Universal Robots URScript: PgProg.script

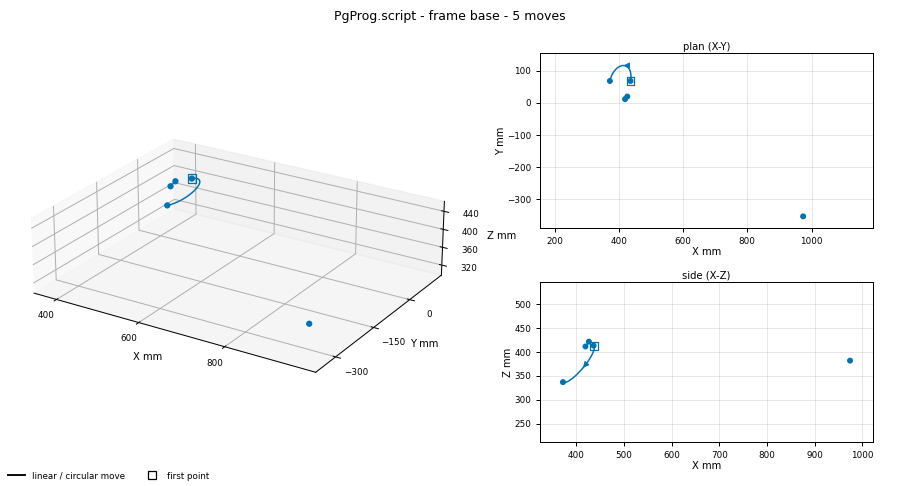
[picture p0: tool path of PgProg.script in frame base, 5 of 9 moves have a stored position in this frame; points joined in program order, loops and branches not executed]
def PgProg():
  # Global parameters:
  global speed_ms    = 0.250
  global speed_rads  = 0.750
  global accel_mss   = 1.200
  global accel_radss = 1.200
  global blend_radius_m = 0.000

  #--------------------------
  # Add any default subprograms here
  # For example, to drive a gripper as a program call:
  # def Gripper_Open():
  #   ...
  # end
  #
  # Example to drive a spray gun:
  def SprayOn(value):
    # use the value as an output:
    DO_SPRAY = 5
    if value == 0:
      set_standard_digital_out(DO_SPRAY, False)
    else:
      set_standard_digital_out(DO_SPRAY, True)
    end
  end

  # Example to synchronize 2
  def Synchronize():
    # Use the following digital output to signal the state of the robot:
    DO_SYNC = 1

    # Use the following digital input to get the state of another robot:
    DI_SYNC = 1

    if (get_standard_digital_out(DO_SYNC) == get_standard_digital_in(DI_SYNC)):
      set_standard_digital_out(DO_SYNC, not (get_standard_digital_out(DI_SYNC)))
      sleep(0.1)
      thread Thread_wait_1():
        while (True):
          sleep(0.01)
        end
      end
      if (get_standard_digital_out(DO_SYNC) != get_standard_digital_in(DI_SYNC)):
        global thread_handler_1=run Thread_wait_1()
        while (get_standard_digital_out(DO_SYNC) != get_standard_digital_in(DI_SYNC)):
          sync()
        end
        kill thread_handler_1
      end
    else:
      if (get_standard_digital_out(DO_SYNC) != get_standard_digital_in(DI_SYNC)):
        set_standard_digital_out(DO_SYNC, not (get_standard_digital_out(DO_SYNC)))
      end
    end
  end

  #
  # Example to move an external axis
  def MoveAxis(value):
    # use the value as an output:
    DO_AXIS_1 = 1
    DI_AXIS_1 = 1
    if value <= 0:
      set_standard_digital_out(DO_AXIS_1, False)

      # Wait for digital input to change state
      #while (get_standard_digital_in(DI_AXIS_1) != False):
      #  sync()
      #end
    else:
      set_standard_digital_out(DO_AXIS_1, True)

      # Wait for digital input to change state
      #while (get_standard_digital_in(DI_AXIS_1) != True):
      #  sync()
      #end
    end
  end
  #--------------------------


  # Main program:
  # Program generated by RoboDK v6.0.7 for ABB IRB 120-3/0.6 on XX/XX/XXXX 18:00:00
  # Using nominal kinematics.
  # Using Ref. Frame Pg: p[1.234570, -0.098765, 0.050500, 0.000000, 0.000000, 0.523599]
  # set_reference(p[1.234570, -0.098765, 0.050500, 0.000000, 0.000000, 0.523599])
  # Using TCP Tool Pg: p[0.010000, 0.020000, 0.150000, 0.261799, 0.000000, 0.000000]
  set_tcp(p[0.010000, 0.020000, 0.150000, 0.261799, 0.000000, 0.000000])
  speed_ms    = 0.2500
  blend_radius_m = 0.0050
  movej([0.000000, -0.174533, 0.349066, 0.000000, 0.523599, 0.000000],1.20000,0.75000,0,0.0000)
  movel(p[0.436232, 0.068297, 0.413715, 0.138328, 2.253250, -0.296646],accel_mss,speed_ms,0,0.005)
  # Circular move (R50.0 mm)
  movec(p[0.414005, 0.116593, 0.367095, 0.138328, 2.253250, -0.296646],p[0.371953, 0.068296, 0.337111, 0.138328, 2.253250, -0.296646],1.20000,0.25000,0.0050)
  movej([0.349066, -0.174533, 0.349066, 0.000000, 0.523599, 0.000000],1.20000,0.75000,0,0.0000)
  accel_radss = 2.094
  speed_rads  = 1.0472
  accel_mss   = 0.8000
  speed_ms    = 0.1000
  movel(p[0.419189, 0.011793, 0.411899, 0.138328, 2.253250, -0.296646],accel_mss,speed_ms,0,0.000)
  blend_radius_m = 0.0000
  movel(p[0.426318, 0.020000, 0.422034, 0.138328, 2.253250, -0.296646],accel_mss,speed_ms,0,0.000)
  sleep(0.500)
  halt() # reimplement this function to force stop
  popup("Hello from postgen","Message",False,False,blocking=True)
  # a comment
  SubProgram()
  CustomCode(42)
  ThreadProg
  set_standard_digital_out(1, True)
  Valve = False
  set_standard_digital_out(3, 2.5)
  while (get_standard_digital_in(2) != True):
    sync()
  end
  while (get_standard_digital_in(4) != False):
    sync()
  end
  # Using TCP Tool2: p[0.000000, 0.000000, 0.200000, 0.000000, 0.000000, 0.000000]
  set_tcp(p[0.000000, 0.000000, 0.200000, 0.000000, 0.000000, 0.000000])
  movej([0.000000, -0.174533, 0.349066, 0.000000, 0.523599, 0.000000],2.09440,1.04720,0,0.0000)
  movej([0.174533, -0.087266, 0.436332, 0.087266, 0.610865, 0.087266],2.09440,1.04720,0,0.0000)
  movel(p[0.973908, -0.353337, 0.382202, -0.503745, 2.359457, 0.000119],accel_mss,speed_ms,0,0.000)
  # End of main program
end

PgProg()
